(* IEC 61131-3 sources: llm-plc-st-eval/data/raw/gpt-4o/I4/zero_shot, 3 files *)

(* ---- ejec_1.st ---- *)
```pascal
FUNCTION_BLOCK FB_EstrellaTriangulo
VAR_INPUT
    btnMarcha : BOOL; // Botón de marcha
    btnParo   : BOOL; // Botón de paro
END_VAR

VAR_OUTPUT
    kM : BOOL := FALSE; // Contactor principal
    kY : BOOL := FALSE; // Contactor estrella
    kD : BOOL := FALSE; // Contactor triángulo
END_VAR

VAR
    estado : INT := 0; // Estado del proceso
    timerEstrella : TON; // Temporizador para el modo estrella
    timerMuerto : TON; // Temporizador para el tiempo muerto
END_VAR

// Inicialización de temporizadores
timerEstrella(IN := FALSE, PT := T#8S);
timerMuerto(IN := FALSE, PT := T#100MS);

IF btnParo THEN
    // Reset de todos los contactores y estado
    kM := FALSE;
    kY := FALSE;
    kD := FALSE;
    estado := 0;
ELSIF btnMarcha THEN
    CASE estado OF
        0: // Estado inicial
            kM := TRUE; // Activar contactor principal
            kY := TRUE; // Activar contactor estrella
            timerEstrella(IN := TRUE); // Iniciar temporizador estrella
            estado := 1; // Cambiar al siguiente estado

        1: // Esperando a que termine el temporizador estrella
            IF timerEstrella.Q THEN
                kY := FALSE; // Desactivar contactor estrella
                timerEstrella(IN := FALSE); // Reset temporizador estrella
                timerMuerto(IN := TRUE); // Iniciar temporizador muerto
                estado := 2; // Cambiar al siguiente estado
            END_IF

        2: // Esperando a que termine el tiempo muerto
            IF timerMuerto.Q THEN
                timerMuerto(IN := FALSE); // Reset temporizador muerto
                kD := TRUE; // Activar contactor triángulo
                estado := 3; // Cambiar al siguiente estado
            END_IF

        3: // Estado final, triángulo activado
            // Mantener kM y kD activados
            // No se requiere acción adicional
    END_CASE
ELSE
    // Si no se presiona btnMarcha, asegurarse de que los contactores están apagados
    kM := FALSE;
    kY := FALSE;
    kD := FALSE;
    estado := 0;
END_IF
END_FUNCTION_BLOCK
```

Este código implementa un arranque estrella-triángulo utilizando un bloque de función en Structured Text (ST) conforme al estándar IEC 61131-3. El bloque maneja el proceso de arranque y parada del motor, asegurando que los contactores estrella y triángulo no estén activos simultáneamente.

(* ---- ejec_2.st ---- *)
```pascal
FUNCTION_BLOCK FB_EstrellaTriangulo
VAR_INPUT
    btnMarcha : BOOL; // Botón de marcha
    btnParo : BOOL;   // Botón de paro
END_VAR

VAR_OUTPUT
    kM : BOOL := FALSE; // Contactor principal
    kY : BOOL := FALSE; // Contactor estrella
    kD : BOOL := FALSE; // Contactor triángulo
END_VAR

VAR
    estado : INT := 0; // Estado del proceso
    timerEstrella : TON; // Temporizador para el tiempo en estrella
    timerMuerto : TON;   // Temporizador para el tiempo muerto
END_VAR

// Inicialización de temporizadores
timerEstrella(IN := FALSE, PT := T#8S);
timerMuerto(IN := FALSE, PT := T#100MS);

IF btnParo THEN
    // Si se presiona el botón de paro, desactivar todos los contactores y reiniciar el estado
    kM := FALSE;
    kY := FALSE;
    kD := FALSE;
    estado := 0;
ELSIF btnMarcha THEN
    CASE estado OF
        0: // Estado inicial
            kM := TRUE; // Activar contactor principal
            kY := TRUE; // Activar contactor estrella
            timerEstrella(IN := TRUE); // Iniciar temporizador de estrella
            estado := 1; // Avanzar al siguiente estado

        1: // Estado de espera en estrella
            IF timerEstrella.Q THEN
                kY := FALSE; // Desactivar contactor estrella
                timerEstrella(IN := FALSE); // Reiniciar temporizador de estrella
                timerMuerto(IN := TRUE); // Iniciar temporizador de tiempo muerto
                estado := 2; // Avanzar al siguiente estado
            END_IF

        2: // Estado de tiempo muerto
            IF timerMuerto.Q THEN
                timerMuerto(IN := FALSE); // Reiniciar temporizador de tiempo muerto
                kD := TRUE; // Activar contactor triángulo
                estado := 3; // Avanzar al siguiente estado
            END_IF

        3: // Estado de operación en triángulo
            // Mantenerse en este estado hasta que se presione el botón de paro
            // No se requiere acción adicional
    END_CASE
ELSE
    // Si no se presiona ningún botón, mantener el estado actual
    // No se requiere acción adicional
END_IF
END_FUNCTION_BLOCK
```

(* ---- ejec_3.st ---- *)
```pascal
FUNCTION_BLOCK FB_EstrellaTriangulo
VAR_INPUT
    btnMarcha : BOOL; // Botón de inicio
    btnParo   : BOOL; // Botón de paro
END_VAR

VAR_OUTPUT
    kM : BOOL := FALSE; // Contactor principal
    kY : BOOL := FALSE; // Contactor estrella
    kD : BOOL := FALSE; // Contactor triángulo
END_VAR

VAR
    timerEstrella : TON; // Temporizador para el modo estrella
    timerMuerto   : TON; // Temporizador para el tiempo muerto
    estado        : INT := 0; // Estado del proceso
END_VAR

// Implementación del arranque estrella-triángulo
IF btnParo THEN
    // Si se presiona el botón de paro, desactivar todos los contactores y reiniciar el estado
    kM := FALSE;
    kY := FALSE;
    kD := FALSE;
    estado := 0;
ELSIF btnMarcha THEN
    CASE estado OF
        0: // Estado inicial
            kM := TRUE; // Activar contactor principal
            kY := TRUE; // Activar contactor estrella
            timerEstrella(IN := TRUE, PT := T#8S); // Iniciar temporizador estrella
            estado := 1; // Cambiar al siguiente estado

        1: // Esperar a que termine el temporizador estrella
            IF timerEstrella.Q THEN
                kY := FALSE; // Desactivar contactor estrella
                timerMuerto(IN := TRUE, PT := T#100MS); // Iniciar temporizador de tiempo muerto
                estado := 2; // Cambiar al siguiente estado
            END_IF

        2: // Esperar a que termine el tiempo muerto
            IF timerMuerto.Q THEN
                kD := TRUE; // Activar contactor triángulo
                estado := 3; // Cambiar al estado final
            END_IF

        3: // Estado final, mantener contactor triángulo activado
            // No se realiza ninguna acción adicional
    END_CASE
ELSE
    // Si no se presiona ningún botón, mantener el estado actual
    timerEstrella(IN := FALSE); // Asegurarse de que el temporizador estrella esté desactivado
    timerMuerto(IN := FALSE); // Asegurarse de que el temporizador muerto esté desactivado
END_IF
END_FUNCTION_BLOCK
```

Este código implementa un arranque estrella-triángulo utilizando un bloque de función en Structured Text (ST) conforme al estándar IEC 61131-3. Se utilizan temporizadores para gestionar los tiempos de conmutación entre los contactores estrella y triángulo, asegurando que nunca estén activos simultáneamente.
